(* IEC 61131-3 sources: open62541_dart/test/plc/plc_programs/schneider_m262, 3 files *)

(* ---- DUT_TestStruct.st ---- *)
// DUT for the OPC UA test fixture struct (M262 / EcoStruxure Machine Expert).
//
// The M262 OPC UA server CAN publish structured data types, so TestStruct is
// present on this controller (supportsComplexTypes = true).
//
// The OPC UA BrowseName of the *instance* is "TestStruct" (declared in
// GVL_Test). Field names + scalar types must match what the tests expect,
// resolved by BrowseName:
//   Id      : DINT   -> OPC UA Int32
//   Value   : REAL   -> OPC UA Float
//   Enabled : BOOL   -> OPC UA Boolean
//   Label   : STRING -> OPC UA String
//
// Create this as a DUT object named "ST_TestStruct" in Machine Expert.
TYPE ST_TestStruct :
STRUCT
    Id      : DINT;
    Value   : REAL;
    Enabled : BOOL;
    Label   : STRING;
END_STRUCT
END_TYPE

(* ---- GVL_Test.st ---- *)
// GVL_Test — OPC UA test fixture for Modicon M262 (EcoStruxure Machine Expert).
// FULL fixture INCLUDING the TestStruct DUT: the M262 OPC UA server supports
// structured data types (matches supportsComplexTypes = true).
//
// Mirrors test/plc/plc_fixture.dart. BrowseNames and IEC types below MUST NOT
// change; the tests resolve every node by BrowseName.
//
// Publishing is done by selecting these variables in the OPC UA Symbol
// Configuration in Machine Expert (see README.md), not with pragmas.
// Paste this declaration into a Global Variable List named "GVL_Test".
VAR_GLOBAL
    // --- Scalars (read/write) ---------------------------------------------
    TestBool    : BOOL;                 // -> OPC UA Boolean
    TestInt     : INT;                  // 16-bit -> OPC UA Int16
    TestDint    : DINT;                 // 32-bit -> OPC UA Int32
    TestReal    : REAL;                 // float32 -> OPC UA Float
    TestLreal   : LREAL;                // float64 -> OPC UA Double
    TestString  : STRING;               // -> OPC UA String

    // --- Writable setpoint (REAL) -----------------------------------------
    Setpoint    : REAL;

    // --- Free-running liveness counter (DINT) -----------------------------
    // Incremented by PLC_PRG every cycle. Read-only from a client's view.
    Counter     : DINT;

    // --- Array[0..9] OF DINT (read/write) ---------------------------------
    TestArray   : ARRAY[0..9] OF DINT;

    // --- Struct instance (read/write) -------------------------------------
    // Published as an OPC UA structured type (Id/Value/Enabled/Label members).
    TestStruct  : ST_TestStruct;
END_VAR

(* ---- PLC_PRG.st ---- *)
// PLC_PRG — cyclic program for the M262 fixture.
// Assign this POU to a cyclic task (e.g. MAST) so Counter actually increments.
//
// Declaration part:
PROGRAM PLC_PRG
VAR
    bInit : BOOL := TRUE;
END_VAR

// Implementation part:
IF bInit THEN
    bInit := FALSE;
    GVL_Test.TestBool   := FALSE;
    GVL_Test.TestInt    := 0;
    GVL_Test.TestDint   := 0;
    GVL_Test.TestReal   := 0.0;
    GVL_Test.TestLreal  := 0.0;
    GVL_Test.TestString := '';
    GVL_Test.Setpoint   := 0.0;
    GVL_Test.Counter    := 0;
    GVL_Test.TestStruct.Id      := 0;
    GVL_Test.TestStruct.Value   := 0.0;
    GVL_Test.TestStruct.Enabled := FALSE;
    GVL_Test.TestStruct.Label   := '';
END_IF

// Liveness counter: increment every scan so clients can prove the program is
// running and measure read/subscription update timing. Wraps at the DINT limit.
GVL_Test.Counter := GVL_Test.Counter + 1;
